// TIA Portal V20 export
// export: Created 2026-10-19T18:38:33.4052814Z, ExportSetting WithDefaults, DisplayName Totally Integrated Automation Portal, DisplayVersion V20 Update 6, DisplayName TIA Portal Openness, DisplayVersion V20 Update 6, DisplayName TIA Portal Version Control Interface, DisplayVersion V20 Update 6, DisplayName SINAMICS Startdrive Advanced, DisplayVersion V20 SP1, DisplayName SINAMICS Startdrive G130, G150, S120, S150, SINAMICS MV, G220, S200, S210, DisplayVersion V20 SP1, DisplayName SINAMICS Startdrive G110M, G120, G120C, G120D, G120P, G115D, DisplayVersion V20 SP1, DisplayName STEP 7 Professional, DisplayVersion V20 Update 6, DisplayName STEP 7 Safety, DisplayVersion V20 Update 2, DisplayName WinCC Basic/Comfort/Advanced, DisplayVersion V20 Update 6, DisplayName WinCC Unified, DisplayVersion V20 Update 6
DATA_BLOCK "Light_Bars_DB_1"   // DB235
VERSION : 0.1
// stored: AutoNumber true, DBAccessibleFromOPCUA true, InstanceOfName Light_Bars, InstanceOfType FB
"Light_Bars"
   // VAR_INPUT
   //    VTD_Mode : UInt;
   //    VTD_Speed : Int;
   //    Fault : Bool;
   // END_VAR
   // VAR_OUTPUT
   //    Animation_B1 : Byte;
   //    Color_B1 : Byte;
   //    Speed_B1 : Byte;
   //    Animation_B2 : Byte;
   //    Color_B2 : Byte;
   //    Speed_B2 : Byte;
   // END_VAR
BEGIN
END_DATA_BLOCK
